INTERFACE I_Status

PROPERTY Running : BOOL
GET
END_GET
END_PROPERTY

PROPERTY Alarm : STRING(80)
GET
END_GET
END_PROPERTY

PROPERTY ProductCount : DINT
GET
END_GET
END_PROPERTY

PROPERTY ActualSpeed : REAL
GET
END_GET
END_PROPERTY

PROPERTY SpeedSetpoint : REAL
GET
END_GET
SET
END_SET
END_PROPERTY

END_INTERFACE

(* stored: Version 1.1.0.1, ProductVersion 3.1 *)
